Fanuc KAREL source: kx00008.compact.KL

PROGRAM KX00008
%STACKSIZE=65535
%PRIORITY=65535
%NOLOCKGROUP
VAR
I : INTEGER
J : INTEGER
B : BOOLEAN
F : FILE
S : STRING[80]
P : XYZWPR
BEGIN
ABORT
END KX00008
